(* IEC 61131-3 sources: sis-interlock-demo/tests/POUs/Suites/FB_CauseEffect_Test, 46 files *)

(* ---- CfgBase.method.decl.st ---- *)
// Матрица тестов: 4 причины, 3 следствия, без срабатывания при старте.
//   1 — задержка 2 с, без обхода;   2 — задержка 5 с, обход до 15 мин, снятие после 30 с нормы;
//   3 — без задержки, обход до 10 с, снятие после 2 с нормы; 4 — выключена.
//   Следствие 1 — причины 1, 2 (16#0003); 2 — причина 3 (16#0004); 3 — все (16#000F). CRC посчитан.
METHOD CfgBase : ST_CemCfg
VAR
    stCfg : ST_CemCfg;   // результат
END_VAR

(* ---- CfgCheckDetectsEachRule.method.decl.st ---- *)
// F_CemCheckCfg: каждое правило таблицы 4.3 даёт свой бит; при CEM_CFG_COUNT причины и следствия не
// проверяются, CRC — всегда
METHOD PRIVATE CfgCheckDetectsEachRule
VAR
    stCfg : ST_CemCfg;      // проверяемая конфигурация
    uBad  : U_SisEnumInt;   // значение вне перечисления
END_VAR

(* ---- CfgErrorRecoveredNeedsReset.method.decl.st ---- *)
// Ошибка конфигурации снята (CfgOk): следствия остаются обесточенными до сброса, первопричина CFG;
// сброс — под напряжением, первопричины нет
METHOD PRIVATE CfgErrorRecoveredNeedsReset
VAR
    fbRig : FB_CemRig;   // стенд
END_VAR

(* ---- CmdBitsCleared.method.decl.st ---- *)
// Импульсы HMI (сброс, обходы, отмены) ФБ сбрасывает в том же вызове
METHOD PRIVATE CmdBitsCleared
VAR
    fbRig : FB_CemRig;   // стенд
END_VAR

(* ---- CrcMismatchAllTripped.method.decl.st ---- *)
// Ручная правка конфигурации без пересчёта CRC: ошибка CEM_CFG_CRC (только она), все выходы обесточены,
// событие CfgError с кодом ошибки
METHOD PRIVATE CrcMismatchAllTripped
VAR
    fbRig : FB_CemRig;     // стенд
    stEv  : ST_SisEvent;   // событие
END_VAR

(* ---- DefaultCfgAllTripped.method.decl.st ---- *)
// Конфигурация по умолчанию (0 причин): до и после вызова все 16 выходов обесточены, ошибка
// CEM_CFG_COUNT, первопричина SIS_FIRST_OUT_CFG, сброс запрещён
METHOD PRIVATE DefaultCfgAllTripped
VAR
    fbRig  : FB_CemRig;   // стенд
    uiJ    : UINT;        // индекс следствия
    xAnyOn : BOOL;        // хотя бы один выход под напряжением
END_VAR

(* ---- DefaultCfgAllTripped.method.impl.st ---- *)
coUnit.TEST('Cem_DefaultCfg_AllTripped');
AssertTrue(Condition := fbRig.fbCem.xTripped, Message := 'before first call: tripped');
fbRig.Cycle();
fbRig.PressReset();
xAnyOn := FALSE;
FOR uiJ := 1 TO GVL_Const.SIS_EFFECTS_MAX DO
    xAnyOn := xAnyOn OR fbRig.Out(uiEffect := uiJ);
END_FOR
AssertFalse(Condition := xAnyOn, Message := 'default cfg: all outputs de-energized');
AssertTrue(Condition := fbRig.fbCem.xTripped, Message := 'default cfg: tripped');
AssertTrue(Condition := fbRig.fbCem.stSts.xCfgError, Message := 'default cfg: config error');
AssertEquals_WORD(Expected := GVL_Const.CEM_CFG_COUNT,
    Actual := fbRig.fbCem.stSts.wCfgErr AND GVL_Const.CEM_CFG_COUNT, Message := 'default cfg: CEM_CFG_COUNT');
AssertEquals_UINT(Expected := GVL_Const.SIS_FIRST_OUT_CFG, Actual := fbRig.fbCem.stSts.uiFirstOut,
    Message := 'default cfg: first-out CFG');
AssertEquals_WORD(Expected := 16#FFFF, Actual := fbRig.fbCem.stSts.wEffectTripped, Message := 'all effects tripped');
AssertFalse(Condition := fbRig.fbCem.stSts.xResetPermitted, Message := 'reset not permitted');
AssertEquals_UINT(Expected := GVL_Const.SIS_FIRST_OUT_CFG, Actual := fbRig.fbCem.stSts.uiResetBlocker,
    Message := 'reset blocker CFG');
AssertEquals_INT(Expected := TO_INT(E_SisEventKind.ResetDenied), Actual := fbRig.fbLog.KindAt(uiBack := 0),
    Message := 'reset denied');
coUnit.TEST_FINISHED();

(* ---- DelayTripsExactlyAtDelay.method.decl.st ---- *)
// Причина 1 с задержкой 2 с: на t0 + 1,9 с не зафиксирована (остаток 100 мс), на t0 + 2,0 с —
// FirstOut, CauseTrip, следствия 1 и 3 обесточены, метка первопричины t0 + 2 с
METHOD PRIVATE DelayTripsExactlyAtDelay
VAR
    fbRig : FB_CemRig;   // стенд
    ltT0  : LTIME;       // момент появления требования
END_VAR

(* ---- DisabledCauseNeverTrips.method.decl.st ---- *)
// Выключенная причина (xEnable = FALSE) не даёт требования и не фиксируется, хотя есть в маске
METHOD PRIVATE DisabledCauseNeverTrips
VAR
    fbRig : FB_CemRig;   // стенд
END_VAR

(* ---- EffectTripEventCarriesCause.method.decl.st ---- *)
// В EffectTrip — младшая зафиксированная причина из маски следствия; уже сработавшее следствие
// нового события не даёт
METHOD PRIVATE EffectTripEventCarriesCause
VAR
    fbRig : FB_CemRig;     // стенд
    stEv  : ST_SisEvent;   // событие
END_VAR

(* ---- EventsOrderInCall.method.decl.st ---- *)
// Порядок событий в одном вызове (6.9): CauseDemand → OverrideOn → ResetDenied → FirstOut → CauseTrip
// → EffectTrip; внутри вида — по возрастанию индекса; номера подряд, метка одна
METHOD PRIVATE EventsOrderInCall
VAR
    fbRig  : FB_CemRig;     // стенд
    stEv   : ST_SisEvent;   // событие
    stLast : ST_SisEvent;   // последнее событие
    udiSeq : UDINT;         // номер события до вызова
END_VAR

(* ---- FirstOutClearedByReset.method.decl.st ---- *)
// Сброс очищает первопричину, метку и маску; следующее срабатывание — новая первопричина, счётчик 2
METHOD PRIVATE FirstOutClearedByReset
VAR
    fbRig : FB_CemRig;   // стенд
END_VAR

(* ---- FirstOutRecordsEarliest.method.decl.st ---- *)
// Первопричина — причина, зафиксированная первой (3 в t0); причина 1, зафиксированная позже, — только
// в wCauseLatched; метка и маска первопричины не меняются
METHOD PRIVATE FirstOutRecordsEarliest
VAR
    fbRig : FB_CemRig;   // стенд
    ltT0  : LTIME;       // момент первой фиксации
END_VAR

(* ---- FirstOutSimultaneousLowestAndMask.method.decl.st ---- *)
// Причины 1 и 3 фиксируются в одном вызове: первопричина — младшая (1), в маске — обе (D-08);
// события CauseTrip — по возрастанию индекса
METHOD PRIVATE FirstOutSimultaneousLowestAndMask
VAR
    fbRig : FB_CemRig;     // стенд
    stEv  : ST_SisEvent;   // событие
END_VAR

(* ---- FirstOutTimestampFromSource.method.decl.st ---- *)
// Метка первопричины и события — время источника I_TimeSource этого вызова
METHOD PRIVATE FirstOutTimestampFromSource
VAR
    fbRig : FB_CemRig;     // стенд
    stEv  : ST_SisEvent;   // событие
END_VAR

(* ---- LatchHeldAfterClear.method.decl.st ---- *)
// Зафиксированная причина остаётся зафиксированной, когда требование ушло; следствие не восстанавливается
METHOD PRIVATE LatchHeldAfterClear
VAR
    fbRig : FB_CemRig;   // стенд
END_VAR

(* ---- MaskBeyondCountCfgError.method.decl.st ---- *)
// Маска следствия с причиной сверх uiCauseCount, непустая маска неиспользуемого следствия и пустая маска
// используемого — ошибка CEM_CFG_EFFECT (CRC пересчитан)
METHOD PRIVATE MaskBeyondCountCfgError
VAR
    fbRig : FB_CemRig;   // стенд
    stCfg : ST_CemCfg;   // проверяемая конфигурация
END_VAR

(* ---- NoTimeSourceUsesSystemTime.method.decl.st ---- *)
// Без источника времени (itfTime = 0) — встроенный PL.FB_SystemTime: причина без задержки фиксируется,
// метка первопричины не нулевая
METHOD PRIVATE NoTimeSourceUsesSystemTime
VAR
    fbCem     : FB_CauseEffect;                                    // ФБ без источника времени
    stCfg     : ST_CemCfg;                                         // конфигурация
    stCmd     : ST_CemCmd;                                         // команды
    axCauseIn : ARRAY[1..GVL_Const.SIS_CAUSES_MAX] OF BOOL;        // требования
END_VAR

(* ---- OverrideCancelAndRequestRestarts.method.decl.st ---- *)
// Снятие и новый запрос обхода в одном вызове (D-13: продление — явной отменой и новым запросом):
// OverrideOff, затем OverrideOn, и новый обход отсчитывается от этого вызова — полные 10 с
// Требование причины 3 держится, чтобы обход не снялся при норме (6.4): проверяется только срок
METHOD PRIVATE OverrideCancelAndRequestRestarts
VAR
    fbRig : FB_CemRig;   // стенд
END_VAR

(* ---- OverrideCancelRestoresTrip.method.decl.st ---- *)
// Снятие обхода командой при действующем требовании: OverrideOff и фиксация в том же вызове
METHOD PRIVATE OverrideCancelRestoresTrip
VAR
    fbRig : FB_CemRig;   // стенд
END_VAR

(* ---- OverrideChatteringNotCleared.method.decl.st ---- *)
// Дребезг требования под пусковым обходом (6.4, D-20): причина 3 (без задержки, обход 10 с, подтверждение
// нормы 2 с); норма каждый раз короче подтверждения (отсчёт доходит до 1,9 с), затем требование на один
// шаг — подтверждение каждый раз начинается заново, OverrideCleared нет; обход снимает срок
// (OverrideExpired) — верхняя граница, и причина с требованием в этом вызове фиксируется
METHOD PRIVATE OverrideChatteringNotCleared
VAR
    fbRig : FB_CemRig;   // стенд
    uiK   : UINT;        // номер периода дребезга
END_VAR

(* ---- OverrideChatteringNotCleared.method.impl.st ---- *)
coUnit.TEST('Cem_Override_ChatteringNotCleared');
fbRig.stCfg := CfgBase();
fbRig.Cycle();
fbRig.stCmd.wOverrideReq := 16#0004;
fbRig.axCauseIn[3] := TRUE;
fbRig.Step(tStep := T#100MS);                                   // t1: обход причины 3 и требование
// 4 периода по 2,1 с: норма в 20 вызовах (подтверждение доходит до 1,9 с), требование — в одном
FOR uiK := 1 TO 4 DO
    fbRig.axCauseIn[3] := FALSE;
    fbRig.Run(tDuration := T#2S, tStep := T#100MS);
    AssertEquals_TIME(Expected := T#100MS, Actual := fbRig.fbCem.stSts.atOverrideClearRemain[3],
        Message := 'chatter: 100 ms of confirm left');
    fbRig.axCauseIn[3] := TRUE;
    fbRig.Step(tStep := T#100MS);
    AssertEquals_TIME(Expected := T#0S, Actual := fbRig.fbCem.stSts.atOverrideClearRemain[3],
        Message := 'chatter: demand resets confirm');
END_FOR
AssertEquals_WORD(Expected := 16#0004, Actual := fbRig.fbCem.stSts.wOverridden,
    Message := 't1 + 8.4 s: override still active');
AssertEquals_UINT(Expected := 0, Actual := fbRig.fbLog.CountKind(eKind := E_SisEventKind.OverrideCleared),
    Message := 'chatter: never cleared');
fbRig.axCauseIn[3] := FALSE;
fbRig.Run(tDuration := T#1S500MS, tStep := T#100MS);            // t1 + 9,9 с
AssertEquals_WORD(Expected := 16#0004, Actual := fbRig.fbCem.stSts.wOverridden,
    Message := 't1 + 9.9 s: override still active');
AssertEquals_TIME(Expected := T#100MS, Actual := fbRig.fbCem.stSts.atOverrideRemain[3],
    Message := 't1 + 9.9 s: 100 ms of override left');
fbRig.axCauseIn[3] := TRUE;
fbRig.Step(tStep := T#100MS);                                   // t1 + 10 с: срок
AssertEquals_UINT(Expected := 1, Actual := fbRig.fbLog.CountKind(eKind := E_SisEventKind.OverrideExpired),
    Message := 't1 + 10 s: OverrideExpired by max time');
AssertEquals_UINT(Expected := 0, Actual := fbRig.fbLog.CountKind(eKind := E_SisEventKind.OverrideCleared),
    Message := 't1 + 10 s: no OverrideCleared');
AssertEquals_WORD(Expected := 0, Actual := fbRig.fbCem.stSts.wOverridden, Message := 't1 + 10 s: no override');
AssertEquals_WORD(Expected := 16#0004, Actual := fbRig.fbCem.stSts.wCauseLatched,
    Message := 't1 + 10 s: demand at expiry latched');
AssertFalse(Condition := fbRig.Out(uiEffect := 2), Message := 't1 + 10 s: effect 2 tripped');
coUnit.TEST_FINISHED();

(* ---- OverrideClearsExactlyAtConfirm.method.decl.st ---- *)
// Автоснятие пускового обхода при норме (6.4, п. 5; R-12): причина 2 (задержка 5 с, обход 15 мин,
// подтверждение нормы 30 с) активна под обходом; требование ушло в t2 — на t2 + 29,9 с обход ещё
// действует (остаток подтверждения 100 мс), ровно на t2 + 30 с — OverrideCleared, без фиксации (требования
// нет); новое требование фиксируется через полную задержку 5 с от своего появления
METHOD PRIVATE OverrideClearsExactlyAtConfirm
VAR
    fbRig : FB_CemRig;     // стенд
    stEv  : ST_SisEvent;   // событие
END_VAR

(* ---- OverrideDelayRunsDuringOverride.method.decl.st ---- *)
// Задержка причины идёт и во время обхода: через 5 с причина 2 активна, но не зафиксирована; снятие
// обхода фиксирует её сразу, без нового отсчёта задержки
METHOD PRIVATE OverrideDelayRunsDuringOverride
VAR
    fbRig : FB_CemRig;   // стенд
END_VAR

(* ---- OverrideDeniedNotAllowed.method.decl.st ---- *)
// Запрос обхода причины без xOverrideAllowed и выключенной причины — OverrideDenied, обхода нет
METHOD PRIVATE OverrideDeniedNotAllowed
VAR
    fbRig : FB_CemRig;     // стенд
    stEv  : ST_SisEvent;   // событие
END_VAR

(* ---- OverrideDeniedWithoutPermit.method.decl.st ---- *)
// Без ключа разрешения обходов разрешённый обход отклоняется
METHOD PRIVATE OverrideDeniedWithoutPermit
VAR
    fbRig : FB_CemRig;   // стенд
END_VAR

(* ---- OverrideExpiresExactly.method.decl.st ---- *)
// Пусковой обход причины 2 (15 мин) и её требование в одном вызове t1: не фиксируется; на
// t1 + 14 мин 59,9 с обход действует (остаток 100 мс); на t1 + 15 мин — OverrideExpired, FirstOut,
// CauseTrip, EffectTrip в одном вызове (задержка 5 с прошла во время обхода)
METHOD PRIVATE OverrideExpiresExactly
VAR
    fbRig : FB_CemRig;   // стенд
END_VAR

(* ---- OverrideExpiryWinsTieWithConfirm.method.decl.st ---- *)
// Срок и подтверждение нормы заканчиваются в одном вызове (6.4: срок проверяется раньше подтверждения):
// обход причины 3 (10 с, подтверждение 2 с) и требование в t1; норма с t1 + 8 с — подтверждение
// заканчивается ровно на t1 + 10 с, вместе со сроком; обход снят по сроку — OverrideExpired, без
// OverrideCleared; требования нет — фиксации нет
METHOD PRIVATE OverrideExpiryWinsTieWithConfirm
VAR
    fbRig : FB_CemRig;   // стенд
END_VAR

(* ---- OverrideRepeatIgnored.method.decl.st ---- *)
// Повторный запрос действующего обхода игнорируется: событий нет, срок не продлевается (D-13).
// Требование причины держится, чтобы обход не снялся при норме (6.4)
METHOD PRIVATE OverrideRepeatIgnored
VAR
    fbRig    : FB_CemRig;   // стенд
    uiEvents : UINT;        // событий до повторного запроса
END_VAR

(* ---- OverrideReRequestAfterExpiryFullTime.method.decl.st ---- *)
// Новый запрос обхода в вызове сразу после истечения прежнего (6.4, п. 4): обход принимается и
// отсчитывается от этого вызова — полный срок 10 с, в этом же вызове не истекает
// Требование причины 3 держится, чтобы обход не снялся при норме (6.4): проверяется только срок
METHOD PRIVATE OverrideReRequestAfterExpiryFullTime
VAR
    fbRig : FB_CemRig;   // стенд
END_VAR

(* ---- OverrideReRequestRestartsConfirm.method.decl.st ---- *)
// Подтверждение нормы и новый обход (6.4, п. 3; D-13): обход причины 3 без требования отсчитывает
// подтверждение (2 с) от вызова, где принят; повторный запрос действующего обхода его не перезапускает;
// снятие и запрос в одном вызове — полные 2 с заново (без Preset подтверждение продолжилось бы); после
// автоснятия новый запрос в следующем вызове — снова полные 2 с, обход не снимается сразу
METHOD PRIVATE OverrideReRequestRestartsConfirm
VAR
    fbRig : FB_CemRig;   // стенд
END_VAR

(* ---- OverrideStartupMaskAllowedOnly.method.decl.st ---- *)
// Общий пусковой обход ставит обходы только включённым причинам с xOverrideAllowed (2 и 3), без
// событий отказа для остальных
METHOD PRIVATE OverrideStartupMaskAllowedOnly
VAR
    fbRig : FB_CemRig;   // стенд
END_VAR

(* ---- ResetAllowedWhenOverridden.method.decl.st ---- *)
// Требование причины под пусковым обходом сбросу не мешает
METHOD PRIVATE ResetAllowedWhenOverridden
VAR
    fbRig : FB_CemRig;   // стенд
END_VAR

(* ---- ResetDeniedWhilePending.method.decl.st ---- *)
// Сброс запрещён и при требовании, которое ещё не прошло задержку (сырое требование, D-07)
METHOD PRIVATE ResetDeniedWhilePending
VAR
    fbRig : FB_CemRig;   // стенд
END_VAR

(* ---- ResetDeniedWhilePresent.method.decl.st ---- *)
// Сброс при требовании причины: ResetDenied с номером мешающей причины, состояние не меняется
METHOD PRIVATE ResetDeniedWhilePresent
VAR
    fbRig : FB_CemRig;     // стенд
    stEv  : ST_SisEvent;   // событие
END_VAR

(* ---- ResetHwEdgeOnly.method.decl.st ---- *)
// Кнопка «Сброс ПАЗ» действует фронтом: удержание не сбрасывает новое срабатывание, нужно отпустить
// и нажать снова
METHOD PRIVATE ResetHwEdgeOnly
VAR
    fbRig : FB_CemRig;   // стенд
END_VAR

(* ---- ResetHwHeldAtStartIgnored.method.decl.st ---- *)
// Кнопка, зажатая при старте ПЛК, — не фронт: срабатывание при старте не сбрасывается
METHOD PRIVATE ResetHwHeldAtStartIgnored
VAR
    fbRig : FB_CemRig;   // стенд
END_VAR

(* ---- ShortPulseNoTrip.method.decl.st ---- *)
// Требование 1,9 с при задержке 2 с не фиксируется (CauseDemand, CauseClear); новое требование
// отсчитывает задержку заново
METHOD PRIVATE ShortPulseNoTrip
VAR
    fbRig : FB_CemRig;   // стенд
END_VAR

(* ---- StartNotTrippedEnergizedFirstCall.method.decl.st ---- *)
// xStartTripped = FALSE: в первом вызове используемые следствия под напряжением (EffectRestore,
// начальное состояние — «сработало»), неиспользуемые обесточены, первопричины нет
METHOD PRIVATE StartNotTrippedEnergizedFirstCall
VAR
    fbRig : FB_CemRig;   // стенд
END_VAR

(* ---- StartTrippedRequiresReset.method.decl.st ---- *)
// xStartTripped = TRUE: после старта все следствия сработали (StartTrip, затем FirstOut START), пока
// оператор не выполнит сброс
METHOD PRIVATE StartTrippedRequiresReset
VAR
    fbRig : FB_CemRig;     // стенд
    stEv  : ST_SisEvent;   // событие
END_VAR

(* ---- TimeBackwardsDuringConfirmEndsOverride.method.decl.st ---- *)
// «Время назад» во время подтверждения нормы (D-19, 6.4): обход причины 2, требование ушло в t2, до
// автоснятия осталось 10 с; источник времени пошёл назад — TimeFault, обход снят как недостоверный по
// сроку (OverrideExpired, не OverrideCleared), подтверждение сброшено, фиксации нет (требования нет);
// позже OverrideCleared не появляется, а новое требование фиксируется через задержку 5 с
METHOD PRIVATE TimeBackwardsDuringConfirmEndsOverride
VAR
    fbRig : FB_CemRig;   // стенд
    ltT2  : LTIME;       // момент, когда требование ушло
END_VAR

(* ---- TimeBackwardsOverrideEnds.method.decl.st ---- *)
// «Время назад» во время пускового обхода (D-19): срок обхода недостоверен — обход снимается в том же
// вызове (OverrideExpired), и причина, задержка которой прошла под обходом, сразу фиксируется
METHOD PRIVATE TimeBackwardsOverrideEnds
VAR
    fbRig : FB_CemRig;   // стенд
    ltT1  : LTIME;       // момент включения обхода
END_VAR

(* ---- TimeBackwardsPendingDelayTrips.method.decl.st ---- *)
// «Время назад» — неисправность источника времени (D-19): отсчёт задержки недостоверен, и причина
// с идущей задержкой срабатывает в том же вызове; причина без требования не срабатывает; событие
// TimeFault — одно
METHOD PRIVATE TimeBackwardsPendingDelayTrips
VAR
    fbRig : FB_CemRig;   // стенд
    ltT0  : LTIME;       // момент появления требования
END_VAR

(* ---- UnusedEffectsDeenergized.method.decl.st ---- *)
// Следствия с номером больше uiEffectCount всегда обесточены
METHOD PRIVATE UnusedEffectsDeenergized
VAR
    fbRig  : FB_CemRig;   // стенд
    uiJ    : UINT;        // индекс следствия
    xAnyOn : BOOL;        // хотя бы один неиспользуемый выход под напряжением
END_VAR

(* ---- UnusedEffectsDeenergized.method.impl.st ---- *)
coUnit.TEST('Cem_UnusedEffects_Deenergized');
fbRig.stCfg := CfgBase();
fbRig.Cycle();
xAnyOn := FALSE;
FOR uiJ := 4 TO GVL_Const.SIS_EFFECTS_MAX DO
    xAnyOn := xAnyOn OR fbRig.Out(uiEffect := uiJ);
END_FOR
AssertFalse(Condition := xAnyOn, Message := 'effects 4..16 de-energized');
AssertTrue(Condition := fbRig.Out(uiEffect := 3), Message := 'used effect 3 energized');
AssertEquals_WORD(Expected := 0, Actual := fbRig.fbCem.stSts.wEffectTripped, Message := 'unused not in wEffectTripped');
AssertFalse(Condition := fbRig.fbCem.xTripped, Message := 'unused effects do not set xTripped');
coUnit.TEST_FINISHED();

(* ---- ZeroDelaySameCall.method.decl.st ---- *)
// Задержка T#0S: причина фиксируется в том же вызове, где появилось требование
METHOD PRIVATE ZeroDelaySameCall
VAR
    fbRig : FB_CemRig;   // стенд
END_VAR
